// TIA Portal V19 export
TYPE "ST_SAFETY_ZONE"
   STRUCT
      SafetyZone_1 : Bool;
      SafetyZone_2 : Bool;
      SafetyZone_3 : Bool;
      SafetyZone_4 : Bool;
      SafetyZone_5 : Bool;
   END_STRUCT;
END_TYPE
